(* Logix 5000 project; controller CIP_14485201 vendor 1 type 14 code 216 rev 38.11; software revision 38.01; part 6 of 11 *)
(* tags used below, declared in another part *)
   Bit : BOOL[128];   // BIT
   Message_Index : ALIAS FOR Integer[30];   // MESSAGE INDEX REGISITER
   Message_Present : INT[5];   // MESSAGES 1-80 PRESENT BITS
   Message_Seq : DINT[101];   // MESSAGE SEQUENCER ARRAY
   Message_Timer : TIMER[1];   // MESSAGE SEQUENCER CONTROL TIMER
   MOA_Status : DINT[10];   // MAN/OFF/AUTO STATUS
   OpCode_Pin : DINT[5];   // OPCODE PIN ARRAY
   PID2 : PID;   // SUPPLY FLOW PID
   PID_Timer : TIMER[5];   // PID TIMERS
   PV_Message : DINT[3];   // PANELVIEW STATUS MESSAGE
   Recipe : RECIPE[41];   // RECIPES
   Sequencer : CONTROL[4];   // SEQUENCER
   Timer : TIMER[99];   // TIMER
   Timer_Chem1_Pump : TIMER[7];   // CHEM #1 CONTROL TIMERS
   Timer_Chem2_Pump : TIMER[7];   // CHEM #2 CONTROL TIMERS
(* MainProgram, continued *)

ROUTINE _06_MESSAGES   (* ladder *)
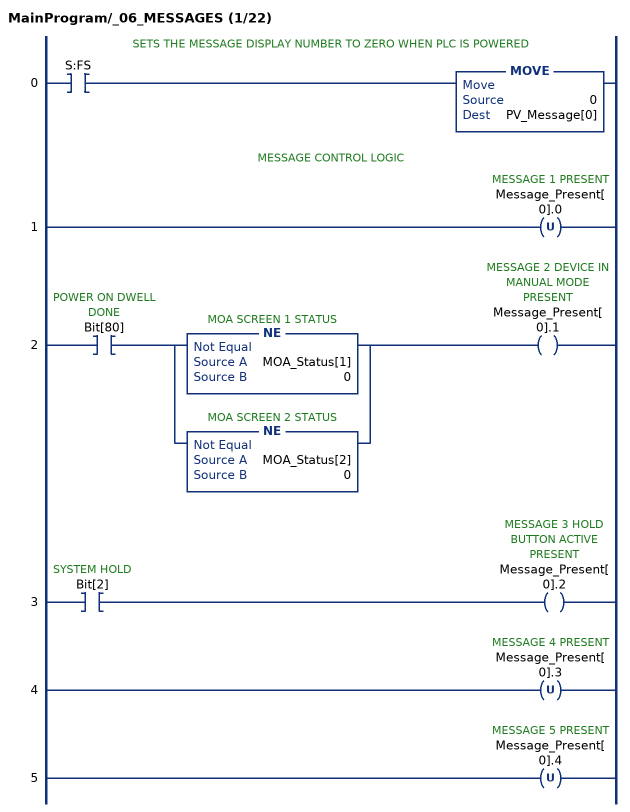
   // SETS THE MESSAGE DISPLAY NUMBER TO ZERO WHEN PLC IS POWERED
   0: XIC(S:FS)MOVE(0,PV_Message[0]);
   // MESSAGE CONTROL LOGIC
   1: OTU(Message_Present[0].0);
   2: XIC(Bit[80])[NE(MOA_Status[1],0) ,NE(MOA_Status[2],0) ]OTE(Message_Present[0].1);
   3: XIC(Bit[2])OTE(Message_Present[0].2);
   4: OTU(Message_Present[0].3);
   5: OTU(Message_Present[0].4);
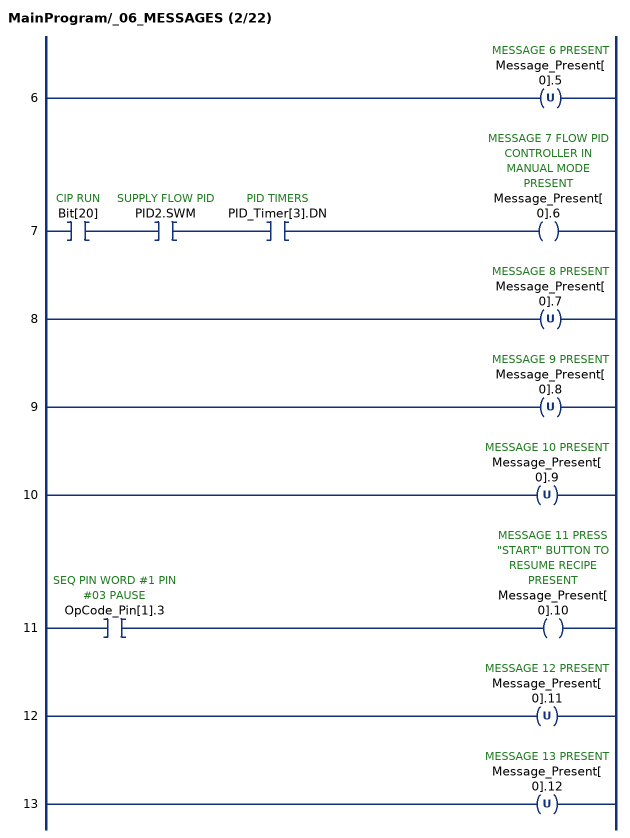
   6: OTU(Message_Present[0].5);
   7: XIC(Bit[20])XIC(PID2.SWM)XIC(PID_Timer[3].DN)OTE(Message_Present[0].6);
   8: OTU(Message_Present[0].7);
   9: OTU(Message_Present[0].8);
   10: OTU(Message_Present[0].9);
   11: XIC(OpCode_Pin[1].3)OTE(Message_Present[0].10);
   12: OTU(Message_Present[0].11);
   13: OTU(Message_Present[0].12);
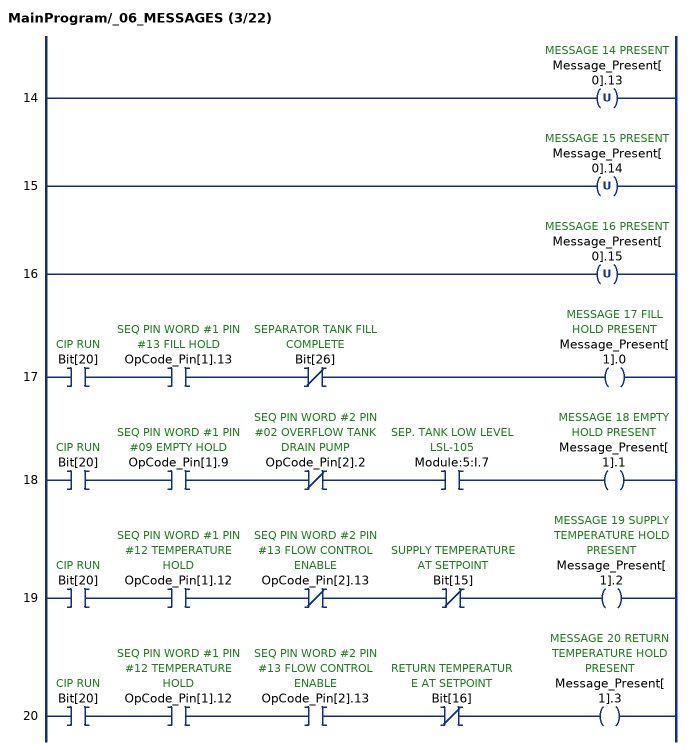
   14: OTU(Message_Present[0].13);
   15: OTU(Message_Present[0].14);
   16: OTU(Message_Present[0].15);
   17: XIC(Bit[20])XIC(OpCode_Pin[1].13)XIO(Bit[26])OTE(Message_Present[1].0);
   18: XIC(Bit[20])XIC(OpCode_Pin[1].9)XIO(OpCode_Pin[2].2)XIC(Module:5:I.7)OTE(Message_Present[1].1);
   19: XIC(Bit[20])XIC(OpCode_Pin[1].12)XIO(OpCode_Pin[2].13)XIO(Bit[15])OTE(Message_Present[1].2);
   20: XIC(Bit[20])XIC(OpCode_Pin[1].12)XIC(OpCode_Pin[2].13)XIO(Bit[16])OTE(Message_Present[1].3);
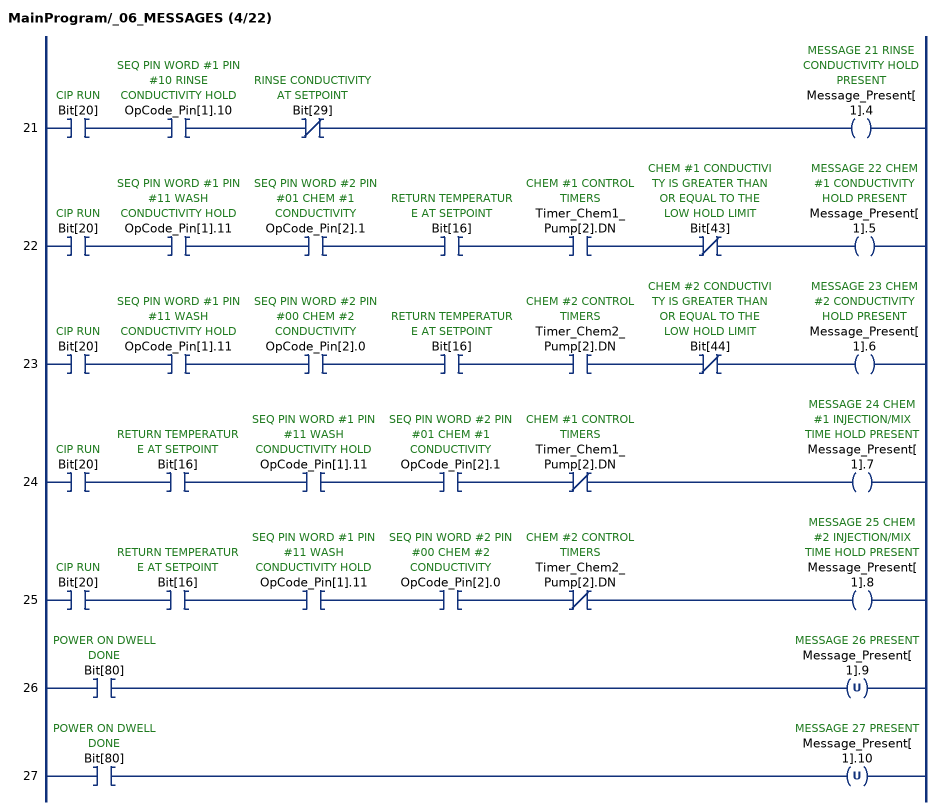
   21: XIC(Bit[20])XIC(OpCode_Pin[1].10)XIO(Bit[29])OTE(Message_Present[1].4);
   22: XIC(Bit[20])XIC(OpCode_Pin[1].11)XIC(OpCode_Pin[2].1)XIC(Bit[16])XIC(Timer_Chem1_Pump[2].DN)XIO(Bit[43])OTE(Message_Present[1].5);
   23: XIC(Bit[20])XIC(OpCode_Pin[1].11)XIC(OpCode_Pin[2].0)XIC(Bit[16])XIC(Timer_Chem2_Pump[2].DN)XIO(Bit[44])OTE(Message_Present[1].6);
   24: XIC(Bit[20])XIC(Bit[16])XIC(OpCode_Pin[1].11)XIC(OpCode_Pin[2].1)XIO(Timer_Chem1_Pump[2].DN)OTE(Message_Present[1].7);
   25: XIC(Bit[20])XIC(Bit[16])XIC(OpCode_Pin[1].11)XIC(OpCode_Pin[2].0)XIO(Timer_Chem2_Pump[2].DN)OTE(Message_Present[1].8);
   26: XIC(Bit[80])OTU(Message_Present[1].9);
   27: XIC(Bit[80])OTU(Message_Present[1].10);
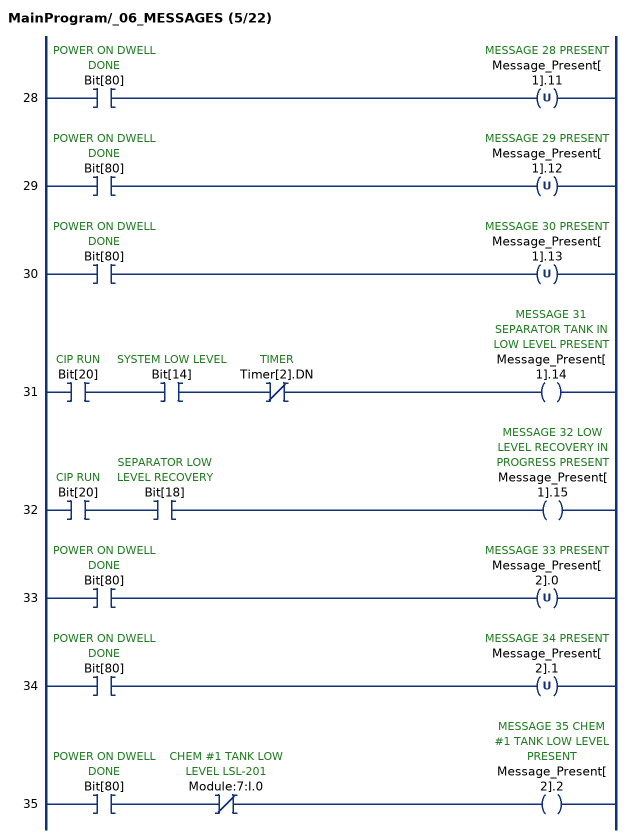
   28: XIC(Bit[80])OTU(Message_Present[1].11);
   29: XIC(Bit[80])OTU(Message_Present[1].12);
   30: XIC(Bit[80])OTU(Message_Present[1].13);
   31: XIC(Bit[20])XIC(Bit[14])XIO(Timer[2].DN)OTE(Message_Present[1].14);
   32: XIC(Bit[20])XIC(Bit[18])OTE(Message_Present[1].15);
   33: XIC(Bit[80])OTU(Message_Present[2].0);
   34: XIC(Bit[80])OTU(Message_Present[2].1);
   35: XIC(Bit[80])XIO(Module:7:I.0)OTE(Message_Present[2].2);
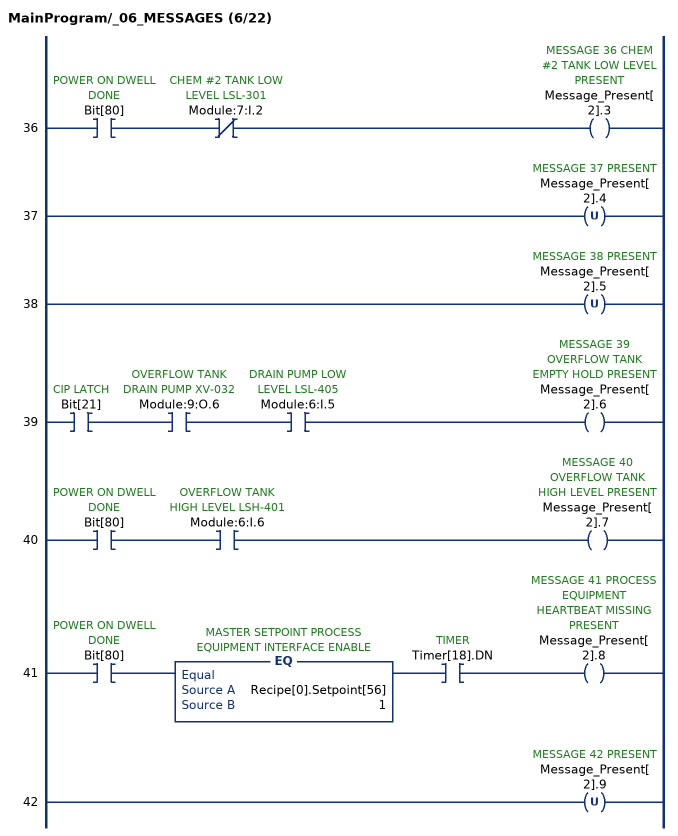
   36: XIC(Bit[80])XIO(Module:7:I.2)OTE(Message_Present[2].3);
   37: OTU(Message_Present[2].4);
   38: OTU(Message_Present[2].5);
   39: XIC(Bit[21])XIC(Module:9:O.6)XIC(Module:6:I.5)OTE(Message_Present[2].6);
   40: XIC(Bit[80])XIC(Module:6:I.6)OTE(Message_Present[2].7);
   41: XIC(Bit[80])EQ(Recipe[0].Setpoint[56],1)XIC(Timer[18].DN)OTE(Message_Present[2].8);
   42: OTU(Message_Present[2].9);
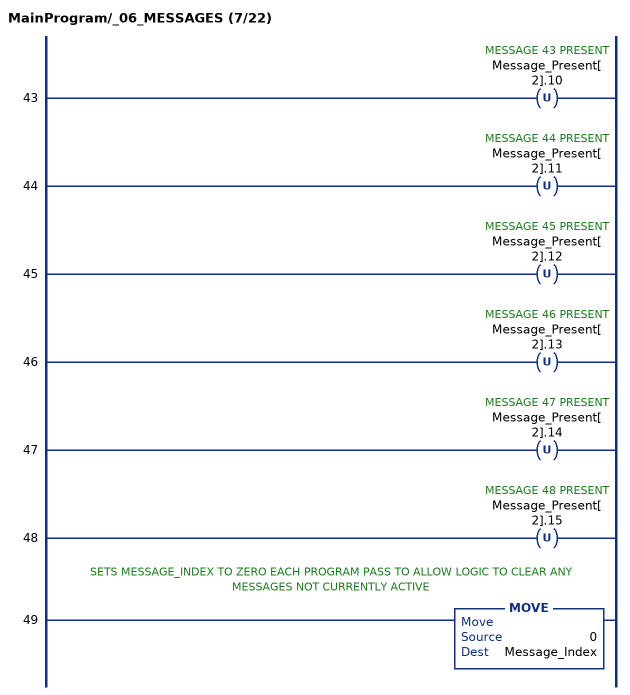
   43: OTU(Message_Present[2].10);
   44: OTU(Message_Present[2].11);
   45: OTU(Message_Present[2].12);
   46: OTU(Message_Present[2].13);
   47: OTU(Message_Present[2].14);
   48: OTU(Message_Present[2].15);
   // SETS MESSAGE_INDEX TO ZERO EACH PROGRAM PASS TO ALLOW LOGIC TO CLEAR ANY MESSAGES NOT CURRENTLY ACTIVE
   49: MOVE(0,Message_Index);
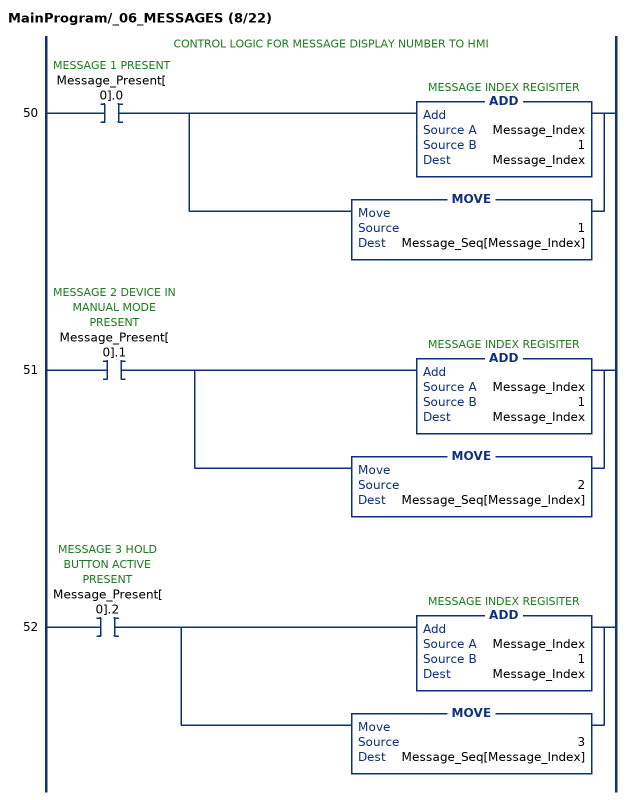
   // CONTROL LOGIC FOR MESSAGE DISPLAY NUMBER TO HMI
   50: XIC(Message_Present[0].0)[ADD(Message_Index,1,Message_Index) ,MOVE(1,Message_Seq[Message_Index]) ];
   51: XIC(Message_Present[0].1)[ADD(Message_Index,1,Message_Index) ,MOVE(2,Message_Seq[Message_Index]) ];
   52: XIC(Message_Present[0].2)[ADD(Message_Index,1,Message_Index) ,MOVE(3,Message_Seq[Message_Index]) ];
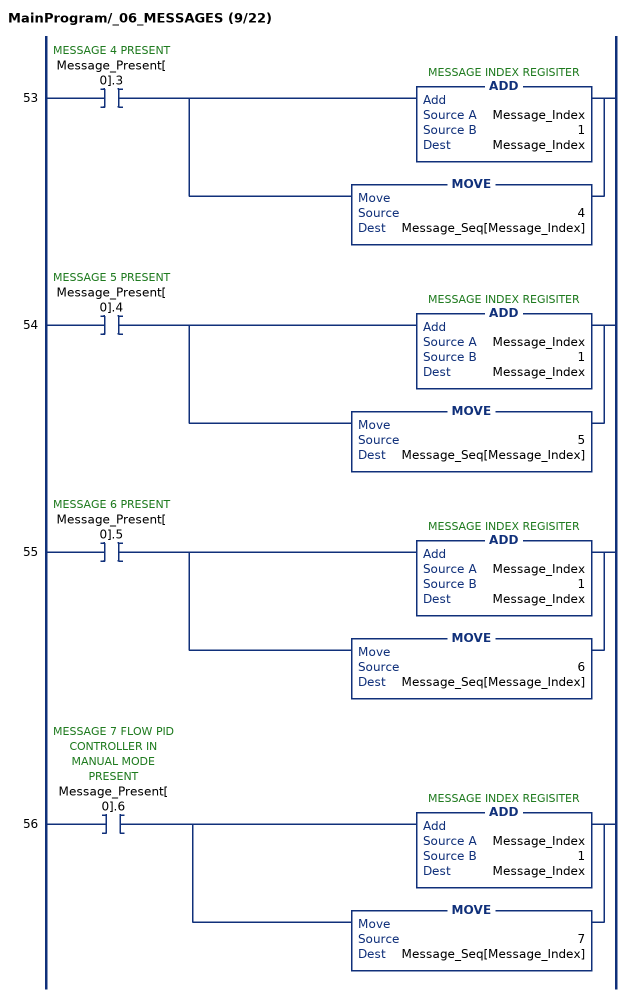
   53: XIC(Message_Present[0].3)[ADD(Message_Index,1,Message_Index) ,MOVE(4,Message_Seq[Message_Index]) ];
   54: XIC(Message_Present[0].4)[ADD(Message_Index,1,Message_Index) ,MOVE(5,Message_Seq[Message_Index]) ];
   55: XIC(Message_Present[0].5)[ADD(Message_Index,1,Message_Index) ,MOVE(6,Message_Seq[Message_Index]) ];
   56: XIC(Message_Present[0].6)[ADD(Message_Index,1,Message_Index) ,MOVE(7,Message_Seq[Message_Index]) ];
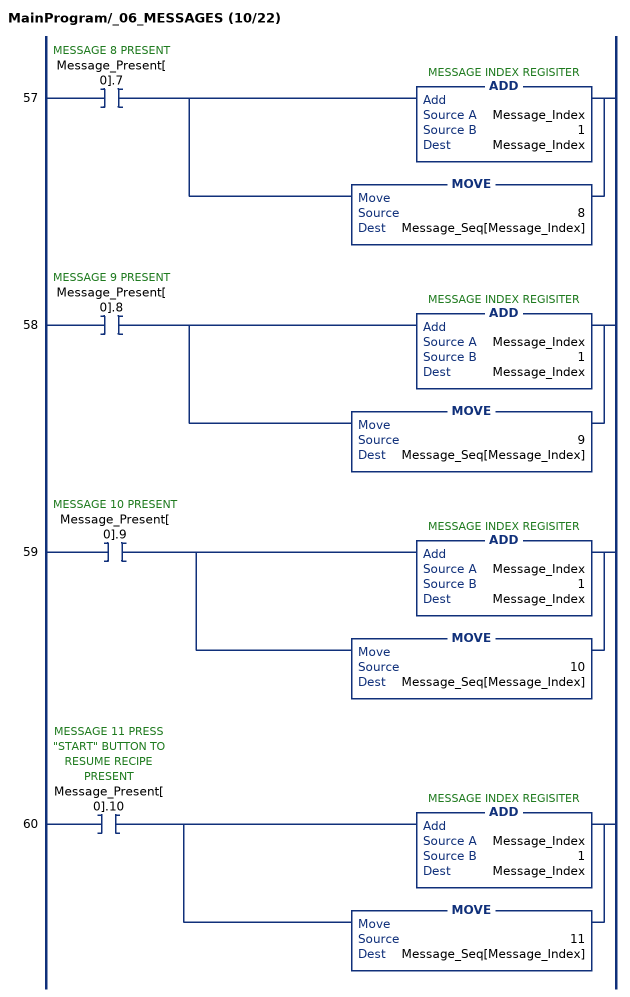
   57: XIC(Message_Present[0].7)[ADD(Message_Index,1,Message_Index) ,MOVE(8,Message_Seq[Message_Index]) ];
   58: XIC(Message_Present[0].8)[ADD(Message_Index,1,Message_Index) ,MOVE(9,Message_Seq[Message_Index]) ];
   59: XIC(Message_Present[0].9)[ADD(Message_Index,1,Message_Index) ,MOVE(10,Message_Seq[Message_Index]) ];
   60: XIC(Message_Present[0].10)[ADD(Message_Index,1,Message_Index) ,MOVE(11,Message_Seq[Message_Index]) ];
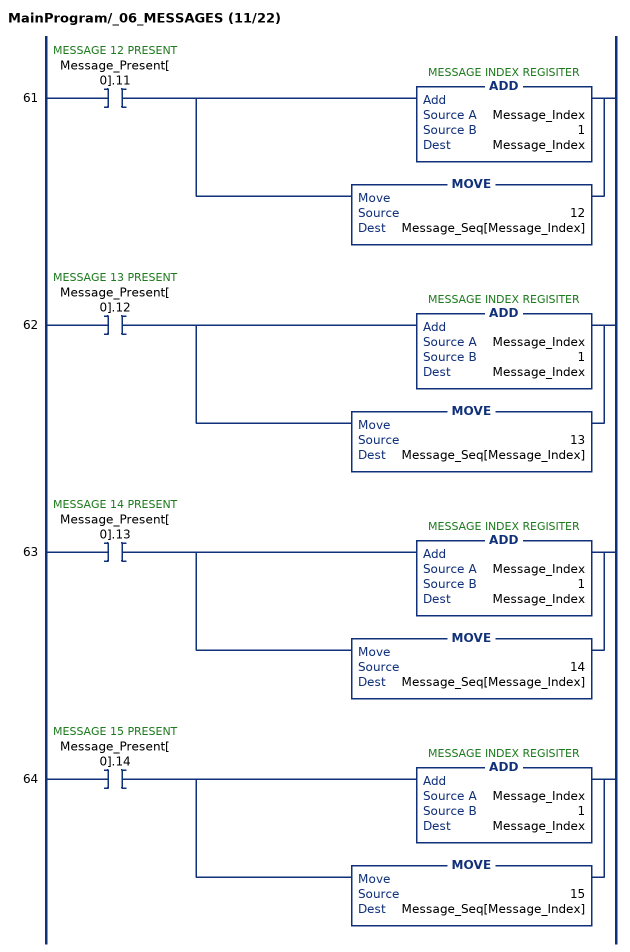
   61: XIC(Message_Present[0].11)[ADD(Message_Index,1,Message_Index) ,MOVE(12,Message_Seq[Message_Index]) ];
   62: XIC(Message_Present[0].12)[ADD(Message_Index,1,Message_Index) ,MOVE(13,Message_Seq[Message_Index]) ];
   63: XIC(Message_Present[0].13)[ADD(Message_Index,1,Message_Index) ,MOVE(14,Message_Seq[Message_Index]) ];
   64: XIC(Message_Present[0].14)[ADD(Message_Index,1,Message_Index) ,MOVE(15,Message_Seq[Message_Index]) ];
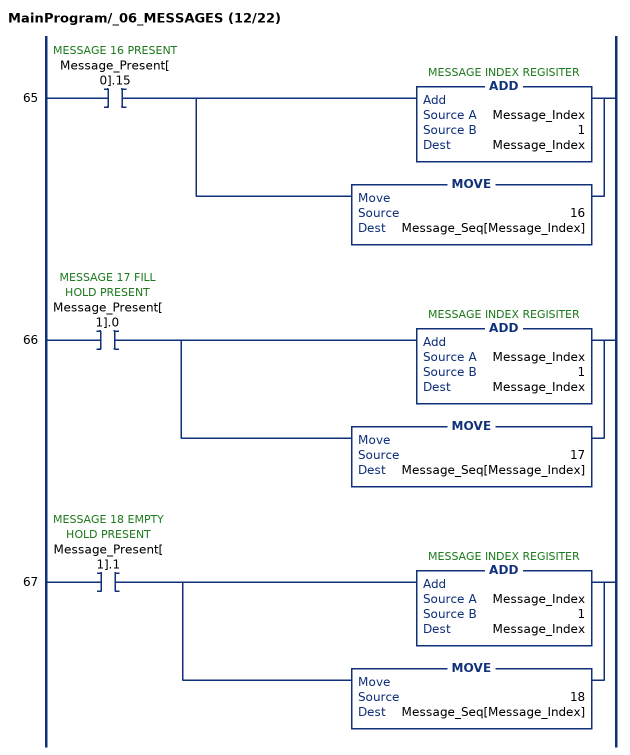
   65: XIC(Message_Present[0].15)[ADD(Message_Index,1,Message_Index) ,MOVE(16,Message_Seq[Message_Index]) ];
   66: XIC(Message_Present[1].0)[ADD(Message_Index,1,Message_Index) ,MOVE(17,Message_Seq[Message_Index]) ];
   67: XIC(Message_Present[1].1)[ADD(Message_Index,1,Message_Index) ,MOVE(18,Message_Seq[Message_Index]) ];
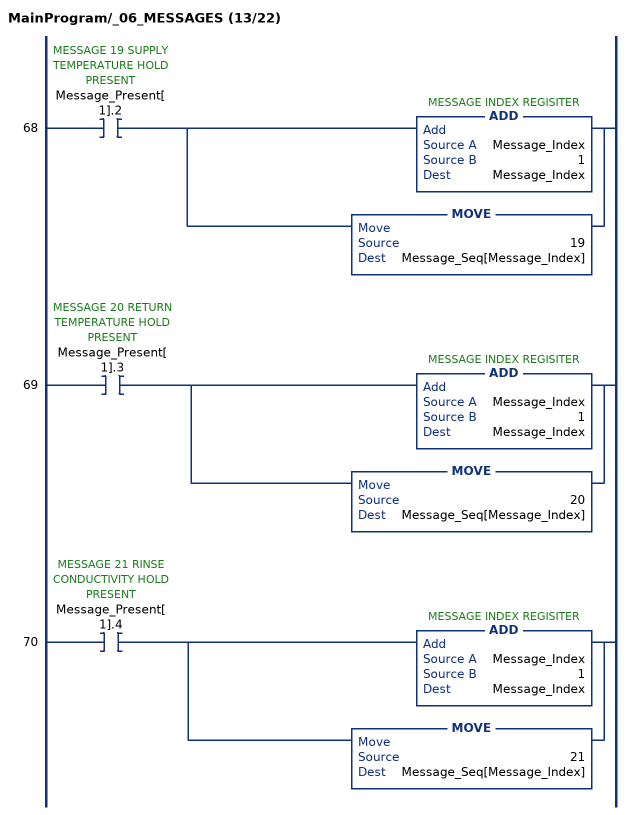
   68: XIC(Message_Present[1].2)[ADD(Message_Index,1,Message_Index) ,MOVE(19,Message_Seq[Message_Index]) ];
   69: XIC(Message_Present[1].3)[ADD(Message_Index,1,Message_Index) ,MOVE(20,Message_Seq[Message_Index]) ];
   70: XIC(Message_Present[1].4)[ADD(Message_Index,1,Message_Index) ,MOVE(21,Message_Seq[Message_Index]) ];
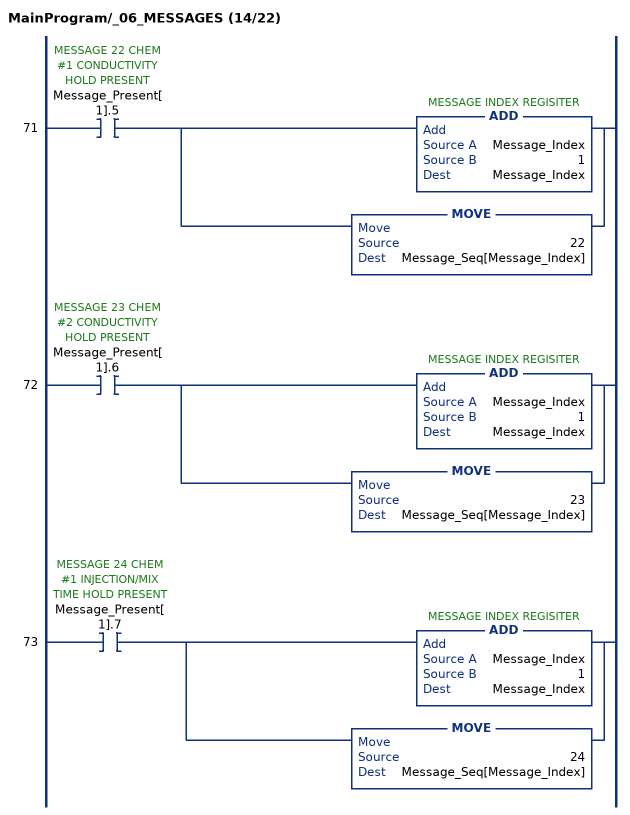
   71: XIC(Message_Present[1].5)[ADD(Message_Index,1,Message_Index) ,MOVE(22,Message_Seq[Message_Index]) ];
   72: XIC(Message_Present[1].6)[ADD(Message_Index,1,Message_Index) ,MOVE(23,Message_Seq[Message_Index]) ];
   73: XIC(Message_Present[1].7)[ADD(Message_Index,1,Message_Index) ,MOVE(24,Message_Seq[Message_Index]) ];
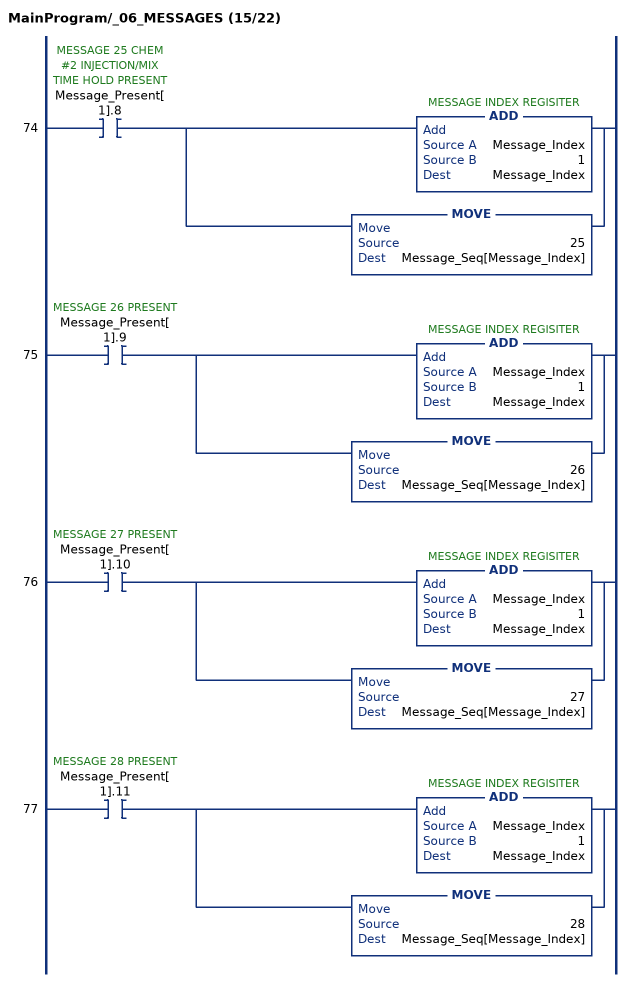
   74: XIC(Message_Present[1].8)[ADD(Message_Index,1,Message_Index) ,MOVE(25,Message_Seq[Message_Index]) ];
   75: XIC(Message_Present[1].9)[ADD(Message_Index,1,Message_Index) ,MOVE(26,Message_Seq[Message_Index]) ];
   76: XIC(Message_Present[1].10)[ADD(Message_Index,1,Message_Index) ,MOVE(27,Message_Seq[Message_Index]) ];
   77: XIC(Message_Present[1].11)[ADD(Message_Index,1,Message_Index) ,MOVE(28,Message_Seq[Message_Index]) ];
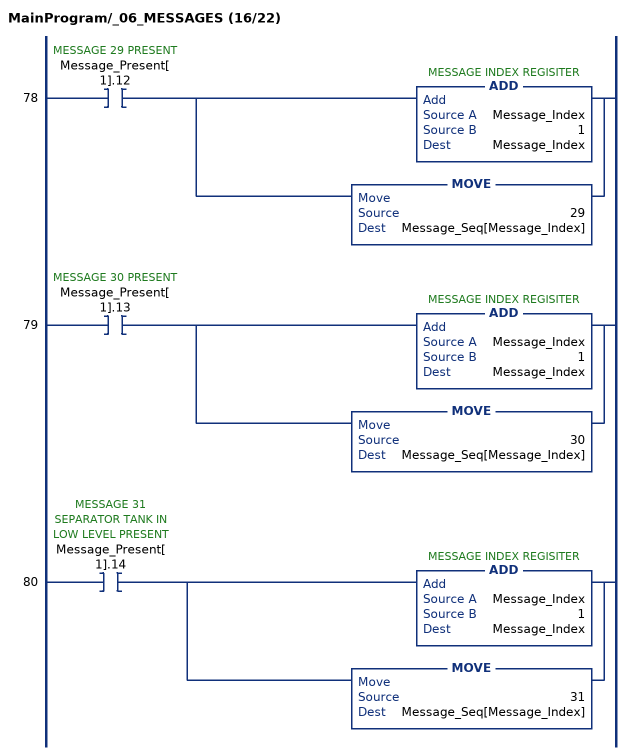
   78: XIC(Message_Present[1].12)[ADD(Message_Index,1,Message_Index) ,MOVE(29,Message_Seq[Message_Index]) ];
   79: XIC(Message_Present[1].13)[ADD(Message_Index,1,Message_Index) ,MOVE(30,Message_Seq[Message_Index]) ];
   80: XIC(Message_Present[1].14)[ADD(Message_Index,1,Message_Index) ,MOVE(31,Message_Seq[Message_Index]) ];
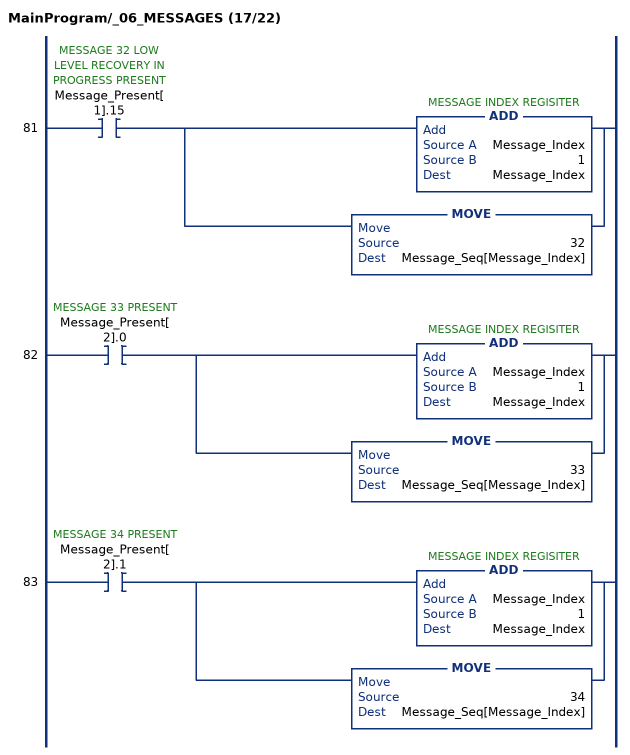
   81: XIC(Message_Present[1].15)[ADD(Message_Index,1,Message_Index) ,MOVE(32,Message_Seq[Message_Index]) ];
   82: XIC(Message_Present[2].0)[ADD(Message_Index,1,Message_Index) ,MOVE(33,Message_Seq[Message_Index]) ];
   83: XIC(Message_Present[2].1)[ADD(Message_Index,1,Message_Index) ,MOVE(34,Message_Seq[Message_Index]) ];
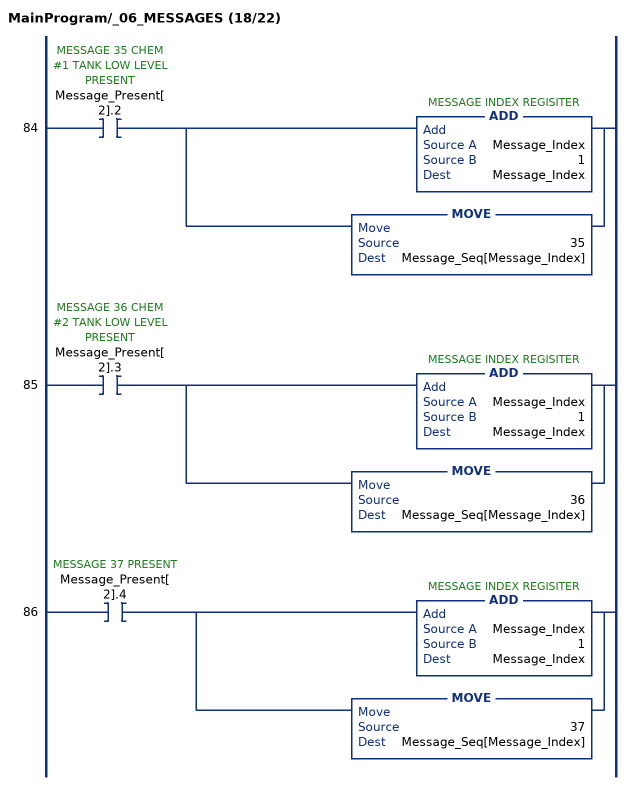
   84: XIC(Message_Present[2].2)[ADD(Message_Index,1,Message_Index) ,MOVE(35,Message_Seq[Message_Index]) ];
   85: XIC(Message_Present[2].3)[ADD(Message_Index,1,Message_Index) ,MOVE(36,Message_Seq[Message_Index]) ];
   86: XIC(Message_Present[2].4)[ADD(Message_Index,1,Message_Index) ,MOVE(37,Message_Seq[Message_Index]) ];
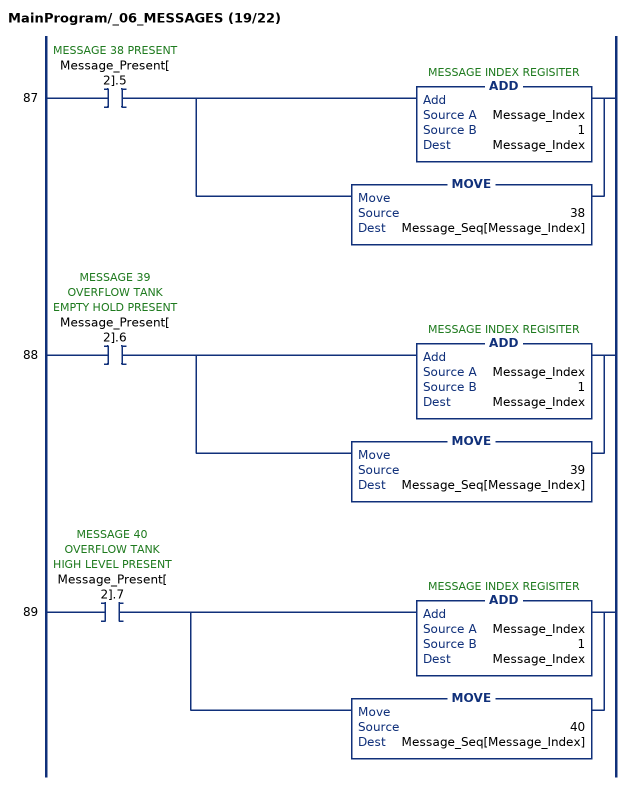
   87: XIC(Message_Present[2].5)[ADD(Message_Index,1,Message_Index) ,MOVE(38,Message_Seq[Message_Index]) ];
   88: XIC(Message_Present[2].6)[ADD(Message_Index,1,Message_Index) ,MOVE(39,Message_Seq[Message_Index]) ];
   89: XIC(Message_Present[2].7)[ADD(Message_Index,1,Message_Index) ,MOVE(40,Message_Seq[Message_Index]) ];
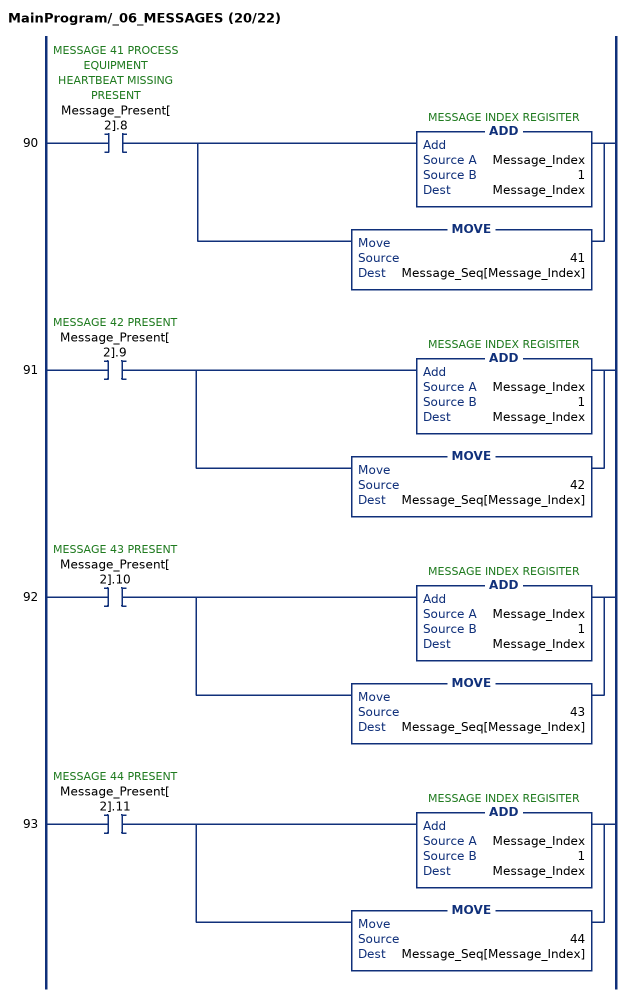
   90: XIC(Message_Present[2].8)[ADD(Message_Index,1,Message_Index) ,MOVE(41,Message_Seq[Message_Index]) ];
   91: XIC(Message_Present[2].9)[ADD(Message_Index,1,Message_Index) ,MOVE(42,Message_Seq[Message_Index]) ];
   92: XIC(Message_Present[2].10)[ADD(Message_Index,1,Message_Index) ,MOVE(43,Message_Seq[Message_Index]) ];
   93: XIC(Message_Present[2].11)[ADD(Message_Index,1,Message_Index) ,MOVE(44,Message_Seq[Message_Index]) ];
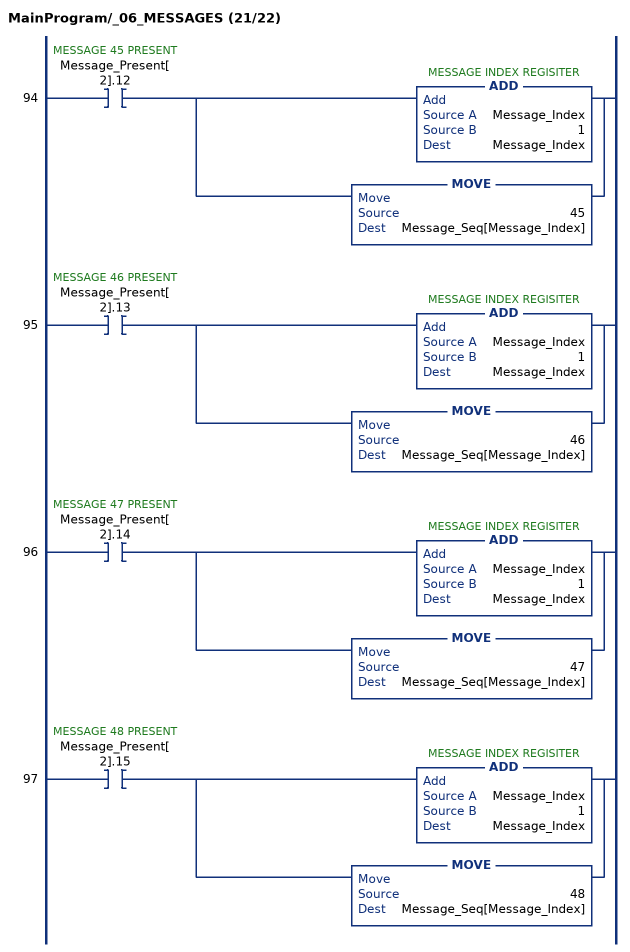
   94: XIC(Message_Present[2].12)[ADD(Message_Index,1,Message_Index) ,MOVE(45,Message_Seq[Message_Index]) ];
   95: XIC(Message_Present[2].13)[ADD(Message_Index,1,Message_Index) ,MOVE(46,Message_Seq[Message_Index]) ];
   96: XIC(Message_Present[2].14)[ADD(Message_Index,1,Message_Index) ,MOVE(47,Message_Seq[Message_Index]) ];
   97: XIC(Message_Present[2].15)[ADD(Message_Index,1,Message_Index) ,MOVE(48,Message_Seq[Message_Index]) ];
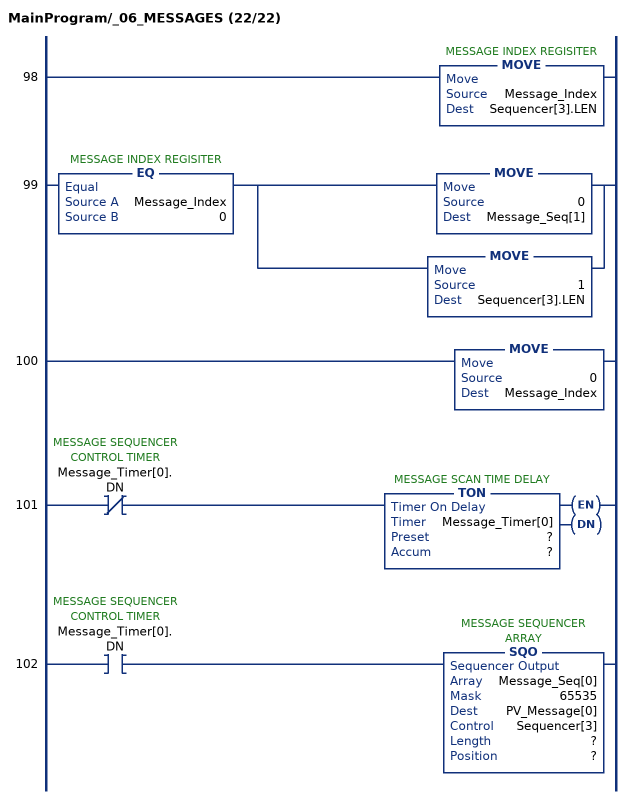
   98: MOVE(Message_Index,Sequencer[3].LEN);
   99: EQ(Message_Index,0)[MOVE(0,Message_Seq[1]) ,MOVE(1,Sequencer[3].LEN) ];
   100: MOVE(0,Message_Index);
   101: XIO(Message_Timer[0].DN)TON(Message_Timer[0],?,?);
   102: XIC(Message_Timer[0].DN)SQO(Message_Seq[0],65535,PV_Message[0],Sequencer[3],?,?);
END_ROUTINE
